Staubli VAL3: plc.pjx

--- plc.pjx ---
Parameters version=s8.21.4cs9_BS4944 stackSize=200000 millimeterUnit=true
Program file=HWcheck.pgx
Program file=changeDataLib.pgx
Program file=changeDataLib1.pgx
Program file=cycle_pause.pgx
Program file=cycle_start.pgx
Program file=cycle_stop.pgx
Program file=init.pgx
Program file=lifebit.pgx
Program file=main.pgx
Program file=powerOnOff.pgx
Program file=receive.pgx
Program file=resetOutput.pgx
Program file=send.pgx
Program file=setSpeed.pgx
Program file=start.pgx
Program file=stop.pgx
Data file=plc.dtx
Library alias=io path=Disk://source/projectSource/io/io.pjx autoload=true password=
Library alias=rs path=Disk://source/projectSource/robotStatus/robotStatus.pjx autoload=true password=
Library alias=savedata path=Disk://source/saveData/saveData.pjx autoload=true password=
Library alias=prog path=Disk://source/projectSource/program/program.pjx autoload=true password=
Library alias=trajectory path=Disk://source/projectSource/trajectory/trajectory.pjx autoload=true password=

--- plc.dtx ---
bool bLifebit = true
bool bReset
bool bSetGun
bool bTosave
public dio dInExcutePainting = {link=3971923C-046E-4FB8-8CDF-8298982DD00B}
dio dInPLCError = {link=0D6C59A5-572E-4845-9D24-D0618D782DD4}
dio dInPowerON = {link=801699AD-0D4E-40AF-A7AF-E7C40311637E}
dio dInResetError = {link=F299EF97-EDDD-4BB8-AA07-719E60051D06}
dio dInStartCycle = {link=842E3CE8-5982-430F-AA8E-B2F701DC178B}
dio dOutCycle = {link=289A5E8D-11F3-4BEB-8FA4-200735E3A2B7}
dio dOutError = {link=79705501-C546-4790-A460-3F340ADFDE5C}
dio dOutEstop = {link=75D4F3C1-C356-4EDA-B423-02C90835EA7D}
dio dOutGunON = {link=734EBAF3-2CA8-4D3F-A8BB-E168C1322725}
dio dOutIsHome = {link=93BF17B5-5C7E-43C6-9C42-3B6025772815}
dio dOutIsPowerd = {link=364EC08F-C077-495B-A954-158507D3C26C}
dio dOutWorkingMode = {link=813E3F4B-A1DE-4C5D-8EAB-0242B6D8A546}
mdesc mNomSpeed
num _bHeavyAlarm
num _nClock = 62473.00582004
num _nNum
num nJointForce[6]
num nLastLib

--- main.pgx ---
public program main()
  local num i
  local bool l_bErr
  local bool l_bLstPower
  local bool l_bValueIn[128]
  local bool l_bValueInLst[128]
  local bool l_bValueOut[128]
  local bool l_bValueOutLst[128]
  local num l_nResult
  local num l_nValue
begin

  call init()
  //call iolink()
  do
    //心跳
    call lifebit()
    //    //硬件检测
    //    call HWcheck()

    //接收信号
    call receive()


    //发送状态
    call send()

    //    //切换数据库
    //    //切换库需要对savedata:nLibIndex做赋值
    //    //库调用函数
    //    //guohangxin modified 20230323
    //    call io:getAnaIO(io:aInput[2],l_nValue,l_bErr)
    //    if workingMode()==4 and l_nValue>0 and l_bErr==false
    //      savedata:nLibIndex=l_nValue
    //      if nLastLib!=savedata:nLibIndex
    //        nLastLib=savedata:nLibIndex
    //        call changeDataLib1(savedata:nLibIndex)
    //        call io:setAnaOutput(io:aOutput[3],savedata:nLibIndex,l_bErr)
    //        //        aioSet(io:aOutput[3],savedata:nLibIndex)
    //        //上位机需要等待发出的lib与收到的反馈lib一致
    //      endIf
    //    else
    //      if nLastLib!=savedata:nLibIndex
    //        nLastLib=savedata:nLibIndex
    //      endIf
    //    endIf
    //    //add by guohangxin 20240408 获取上升沿下降沿信号
    //    for i=0 to size(io:dInput)-1
    //      call io:getDigIO(io:dInput[i],l_bValueIn[i],l_bErr)
    //      if l_bValueIn[i]==true and l_bValueInLst[i]==false
    //        l_bValueInLst[i]=l_bValueIn[i]
    //        rs:sIOStatus="dIn"+toString("",i)+"=ON"
    //      endIf
    //      if l_bValueIn[i]==false and l_bValueInLst[i]==true
    //        l_bValueInLst[i]=l_bValueIn[i]
    //        rs:sIOStatus="dIn"+toString("",i)+"=OFF"
    //      endIf
    //    endFor

    //    for i=0 to size(io:dOutput)-1
    //      //排除掉心跳信号的上升沿下降沿
    //      if i!=7
    //        call io:getDigIO(io:dOutput[i],l_bValueOut[i],l_bErr)
    //        if l_bValueOut[i]==true and l_bValueOutLst[i]==false
    //          l_bValueOutLst[i]=l_bValueOut[i]
    //          rs:sIOStatus="dOut"+toString("",i)+"=ON"
    //        endIf
    //        if l_bValueOut[i]==false and l_bValueOutLst[i]==true
    //          l_bValueOutLst[i]=l_bValueOut[i]
    //          rs:sIOStatus="dOut"+toString("",i)+"=OFF"
    //        endIf
    //      endIf
    //    endFor
    //    //机器人异常检测（碰撞给出信号等）
    //    //如果机器人处于running或held暂停状态，且工作模式未远程自动
    //    //此时如果从上电状态到下点状态，则说明有异常
    //    if(rs:_nOmacStat==3 or rs:_nOmacStat==6) and workingMode()==4 and isPowered()==false and l_bLstPower==true
    //      l_bLstPower=false
    //      //观察1秒钟查看当前工作模式有没有切换，如果有切换，说明认为切换到了手动，此时不做报警处理
    //      if watch(workingMode()!=4,1)==false
    //        call rs:setAlarm(303,0)
    //        call rs:saveLog("",l_nResult)
    //      endIf
    //    elseIf isPowered()==true
    //      l_bLstPower=true
    //    endIf
    delay(0)
  until false
end

--- start.pgx ---
program start()
begin
end

--- changeDataLib.pgx ---
public program changeDataLib(num x_nLib (dimensions=1))
  local num l_nResult
begin
  //形参：x_nLib
  //对应实参：savedata:nLibIndex
  bTosave=true
  call trajectory:onSave(bTosave)
  bTosave=true
  call prog:onSave(bTosave)
  call trajectory:loadTRAJ(x_nLib,l_nResult)
  call prog:loadPROG(x_nLib,l_nResult)

end

--- changeDataLib1.pgx ---
public program changeDataLib1(num x_nLib (dimensions=1))
  local num l_nClock
  local num l_nResult
begin
  //形参：x_nLib
  //对应实参：savedata:nLibIndex
  //  bTosave=true
  //  call trajectory:onSave(bTosave)
  //  bTosave=true
  //  call prog:onSave(bTosave)
  l_nClock=clock()
  logMsg("自动开始切换库:"+toString(".2",clock()))
  call trajectory:loadTRAJ(x_nLib,l_nResult)
  call prog:loadPROG(x_nLib,l_nResult)

  delay(1)
  logMsg(toString(".3",clock()-l_nClock))
end

--- cycle_pause.pgx ---
public program cycle_pause()
begin
  rs:bToPause=true
  //  wait(rs:bIsPause==true)
  //  rs:bToPause=false
  //  logMsg("PLC:pausecycle")
end

--- cycle_start.pgx ---
public program cycle_start()
begin
  rs:bToStartCycle=true
  wait(rs:bIsCycle==true)
  rs:bToStartCycle=false


  logMsg("PLC:startcycle")
end

--- cycle_stop.pgx ---
public program cycle_stop()
begin
  rs:bToStopCycle=true
  stopMove()
  wait(rs:bIsCycle==false)
  rs:bToStopCycle=false
  logMsg("PLC:stopcycle")
end

--- HWcheck.pgx ---
public program HWcheck()
  local num l_nNum
  local num l_nState
  local num l_nState1
  local string l_sState
begin
  //  rs:nHWState=$getState()
  //  l_nState=rs:nHWState
  //  if l_nState<0
  //    if !bReset
  //      l_nState=abs(l_nState)-90
  //      l_nState1=roundDown(l_nState)
  //      switch l_nState1
  //        case 0

  //          call rs:setAlarm(400,0)
  //        break
  //        case 1
  //          l_nNum= aioGet(ainRSI)
  //          if l_nNum!=0
  //            call rs:setAlarm(401,0)
  //          endIf
  //        break
  //        case 2
  //          call rs:setAlarm(402,0)
  //        break
  //        case 3
  //          call rs:setAlarm(403,0)
  //        break
  //        case 4
  //          call rs:setAlarm(404,0)
  //        break
  //        case 5
  //          call rs:setAlarm(405,0)
  //        break

  //      endSwitch
  //      bReset=true
  //    endIf
  //  else
  //    bReset=false
  //  endIf
end

--- init.pgx ---
program init()
begin
  _nClock=0
  call io:init()
end

--- lifebit.pgx ---
public program lifebit()
begin
  //  _nClock=0
  //  do
  if clock()-_nClock>1
    _nClock=clock()
    bLifebit=!bLifebit
  endIf


  //  delay(0)
  //  until false
end

--- powerOnOff.pgx ---
public program powerOnOff(bool x_bPowerOn (dimensions=1))
begin
  if x_bPowerOn==true
    //Power on
    if !isPowered() and esStatus()!=2 and workingMode()==4
      autoConnectMove(true)
      enablePower()
      delay(1)
    endIf
  else
    //Power Off
    if isPowered()
      disablePower()
      delay(1)
    endIf
  endIf
end

--- receive.pgx ---
public program receive()
  local bool l_bAckAlarm
  local bool l_bEndCmd
  local bool l_bErr
  local bool l_bHoldCmd
  local bool l_bPowerOff
  local bool l_bPowerOn
  local bool l_bResetCmd
  local bool l_bResetIO
  local bool l_bResult
  local bool l_bRotToHome
  local bool l_bStartCmd
  local bool l_bStopCmd
  local bool l_bToHome
  local bool l_bValue
  local num l_n
  local num l_nResult
  local num l_nSpeed
begin
  //机器人上电
  if dInPowerON==true and !isPowered() and workingMode()==4 and !rs:bIsEstop
    enablePower()
    l_bResult=watch(isPowered()==true,1)
    if !l_bResult
      popUpMsg("机器人上电超时")
    endIf
  endIf

  if rs:bIsCycle and workingMode()==1
    call cycle_stop()
  endIf
  //启动主程序
  if dInStartCycle==true and !rs:bIsCycle and rs:bIsHome and workingMode()==4 and !rs:bIsEstop
    //复位信号
    // call resetOutput()
    //
    //call cycle_stop()
    resetMotion()
    call cycle_start()
  endIf
  //暂停&恢复
  if dInPLCError==true
    if dOutGunON==true
      bSetGun=true
      dOutGunON=false
    endIf
    if rs:bIsCycle
      call cycle_pause()
    endIf
  elseIf dInPLCError==false and rs:bIsPause
    if bSetGun
      dOutGunON=true
    endIf
    call cycle_start()
  endIf
  //复位报警
  if dInResetError==true
    rs:bIsError=false
  endIf

  //设置速度
  call setSpeed()

  if esStatus()==1
    setSafetyRestart()
  endIf


end

--- resetOutput.pgx ---
public program resetOutput()
  local bool l_bErr
  local num l_nI
begin
  //2025.7.21 add 复位输出信号
  for l_nI=9 to size(io:dOutput)-1
    call io:setDigOutput(io:dOutput[l_nI],false,l_bErr)
  endFor
  for l_nI=0 to size(io:aOutput)-1
    call io:setAnaOutput(io:aOutput[l_nI],0,l_bErr)
  endFor
end

--- send.pgx ---
program send()
  local num i
  local bool l_bEnabling
  local bool l_bErr
  local bool l_bLastPower
  local bool l_bMcpEstop
  local num l_i
begin
  //远程模式
  dOutWorkingMode=rs:bIsRemoteAuto
  //上电
  dOutIsPowerd=isPowered()
  //程序运行
  dOutCycle=rs:bIsCycle
  //机器人报警
  dOutError=rs:bIsError
  //机器人急停
  dOutEstop=rs:bIsEstop
  //机器人在原点
  dOutIsHome=rs:bIsHome
  //机器人通讯故障
  if ioStatus(dOutIsHome)<0
    rs:bIsError=true
  endIf
end

--- send1.pgx ---
program send()
  local num l_i
  local bool l_bErr
  local num i
  local bool l_bMcpEstop
  local bool l_bEnabling
begin

  //状态
  rs:bIsHome=(abs((herej()-savedata:jHome))<{2,2,2,2,2,2})
  rs:bIsEstop=(io:dRSI9["RbStop"]==false)
  rs:bIsReady=(rs:_nOmacStat==1)
  rs:bIsCycle=(rs:_nOmacStat==3)

  call io:setDigOutput(io:dORbAtHome,rs:bIsHome,l_bErr)
  //stop
  call io:setDigOutput(io:dORbStopped,(rs:_nOmacStat==9),l_bErr)
  call io:setDigOutput(io:dORbReady,(rs:_nOmacStat==1),l_bErr)
  call io:setDigOutput(io:dORbRunning,(rs:_nOmacStat==3),l_bErr)
  call io:setDigOutput(io:dORbHeld,(rs:_nOmacStat==6),l_bErr)
  call io:setDigOutput(io:dORbManualMode,(workingMode()==1),l_bErr)
  call io:setDigOutput(io:dORbAutoMode,(workingMode()==4),l_bErr)
  call io:getDigIO(io:dRSI9["enabling"],l_bEnabling,l_bErr)
  call io:setDigOutput(io:dORbEnable,(l_bEnabling==true),l_bErr)
  call io:getDigIO(io:dRSI9["RbStop"],l_bMcpEstop,l_bErr)
  call io:setDigOutput(io:dOMcpEstop,(l_bMcpEstop==false),l_bErr)
  call io:setDigOutput(io:dORbMoving,!isSettled(),l_bErr)
  call io:setDigOutput(io:dORbHeartbeat,bLifebit,l_bErr)
  call io:setDigOutput(io:dORbPowerOn,isPowered(),l_bErr)

  //
  for i=0 to size(rs:_nAlarmCode)-1
    if rs:_nAlarmCode[i]>rs:nHeavyAlarmLev
      rs:_bHeavyAlarm=true
      //1.机器人错误代码
      call io:setAnaOutput(io:aOutput[2],rs:_nAlarmCode[rs:_nErrIndex],l_bErr)
    endIf
  endFor
  if rs:_bHeavyAlarm
    call io:setDigOutNoAlm(io:dORbAlarm,true,l_bErr)
  else
    call io:setDigOutNoAlm(io:dORbAlarm,false,l_bErr)
  endIf
  //  //jointforce
  //  getJointForce(nJointForce)
  //  for l_i = 0 to size(nJointForce)-1
  //    call io:setAnaOutput(io:aOutput[l_i],nJointForce[l_i],l_bErr)
  //  endFor

  //************************模拟量输出*****************************
  //0.机器人当前的运动速度
  call io:setAnaOutput(io:aOutput[1],getMonitorSpeed(),l_bErr)
  //1.反馈程序号
  call io:setAnaOutput(io:aOutput[0],rs:nProgCode,l_bErr)
end

--- setSpeed.pgx ---
program setSpeed()
  local bool l_bErr
  local num l_nResult
  local num l_nSpeed
begin
  //设置机器人速度
  if getProfile()=="customer"
    call io:getAnaIO(io:aInput[1],l_nSpeed,l_bErr)
    if l_bErr==false
      l_nSpeed=round(l_nSpeed)
      if l_nSpeed>0 and l_nSpeed<=100 and getMonitorSpeed()!=l_nSpeed
        setMonitorSpeed(l_nSpeed)
      endIf
    endIf
  endIf
  //手动设回default权限
  if workingMode()==4 and getProfile()!="customer"
    l_nResult=setProfile("customer","")
  endIf
  if workingMode()==1 and getProfile()=="customer"
    l_nResult=setProfile("default","")
  endIf
end

--- stop.pgx ---
program stop()
begin
end
